(* IEC 61131-3 sources: iolistgen/tools/tests/fixtures/lowering/src/GVLs, 1 file *)

(* ---- GVL_Const.gvl.st ---- *)
// Константы примера понижения: границы массивов и длины строк вычисляются по ним
VAR_GLOBAL CONSTANT
    SLOTS_MAX : UINT := 4;
    GRID_MAX : UINT := SLOTS_MAX * 2 - 1;
    NAME_LEN : UINT := 16#20;
END_VAR
